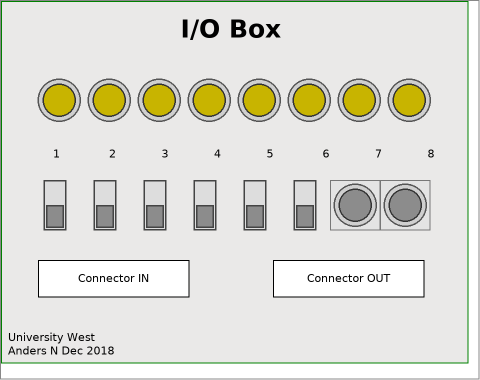
VISUALIZATION Visualization  // 480x380
    Rectangle (1,1 467x362)
    Label (147,0 168x57), "I/O Box"
    Lamp1 (34,75 50x50), variable: GVL.ixLed1, style: Lamp-Lamp1-Yellow
    Lamp1 (84,75 50x50), variable: GVL.ixLed2, style: Lamp-Lamp1-Yellow
    Lamp1 (134,75 50x50), variable: GVL.ixLed3, style: Lamp-Lamp1-Yellow
    Lamp1 (184,75 50x50), variable: GVL.ixLed4, style: Lamp-Lamp1-Yellow
    Lamp1 (234,75 50x50), variable: GVL.ixLed5, style: Lamp-Lamp1-Yellow
    Lamp1 (284,75 50x50), variable: GVL.ixLed6, style: Lamp-Lamp1-Yellow
    Lamp1 (334,75 50x50), variable: GVL.ixLed7, style: Lamp-Lamp1-Yellow
    Lamp1 (384,75 50x50), variable: GVL.ixLed8, style: Lamp-Lamp1-Yellow
    Label (5,329 118x30), "University West Anders N Dec 2018"
    Label (50,144 392x20), "1 2 3 4 5 6 7 8"
    RoundedRectangle (38,260 151x37), "Connector IN"
    RoundedRectangle (273,260 151x37), "Connector OUT"
    DipSwitch (30,180 50x50), variable: GVL.qxButton1, behaviour: TOGGLE, style: Switch-DipSwitch-Gray
    DipSwitch (80,180 50x50), variable: GVL.qxButton2, behaviour: TOGGLE, style: Switch-DipSwitch-Gray
    DipSwitch (130,180 50x50), variable: GVL.qxButton3, behaviour: TOGGLE, style: Switch-DipSwitch-Gray
    DipSwitch (180,180 50x50), variable: GVL.qxButton4, behaviour: TOGGLE, style: Switch-DipSwitch-Gray
    DipSwitch (230,180 50x50), variable: GVL.qxButton5, behaviour: TOGGLE, style: Switch-DipSwitch-Gray
    DipSwitch (280,180 50x50), variable: GVL.qxButton6, behaviour: TOGGLE, style: Switch-DipSwitch-Gray
    PushSwitch (330,180 50x50), variable: GVL.qxButton7, behaviour: TAP, style: Switch-PushSwitch-Gray
    PushSwitch (380,180 50x50), variable: GVL.qxButton8, behaviour: TAP, style: Switch-PushSwitch-Gray
    hotkey HotkeyInput Id=481044725760, Key=KeyName=1, VisuElemId=-1
END_VISUALIZATION

(* stored: Version 1.1.0.1, ProductVersion 3.1.4024.12
   Visu Visualization: Id {f3ed196b-a41c-4cdb-befe-4a966ff196a9} *)
